{attribute 'qualified_only'}
VAR_GLOBAL
    // inputs
    xPressureOK, xEStop                         : BOOL;
    xLS_Infeed, xLS_Outfeed                     : BOOL;
    xServoInLatched, xServoInAS, xServoInGS     : BOOL;
    xServoOutLatched, xServoOutAS, xServoOutGS  : BOOL;
    xCW_Lready, xCW_JobLoaded, xCW_MarkBusy     : BOOL;
    // cylinders (valves = outputs, sensors = inputs)
    stInfeed, stOutfeed, stEjector, stClamp, stDiverter : ST_CylIO;
    // outputs
    xVent, xLaserEnable, xCW_Trig, xCW_STO      : BOOL;
    nCW_Job                                     : USINT;   // job number 0..15
    xBlowAS, xBlowGS, xBypassAS, xBypassGS      : BOOL;
END_VAR

(* stored: Version 1.1.0.1
   GVL GVL_IO: Id {5b15ce66-8e0e-4326-b088-54bac4a0ea54} *)
